// TIA Portal V21 export
FUNCTION_BLOCK "Mixed"   // FB1, LAD
BEGIN

REGION Network 1: Unknown part
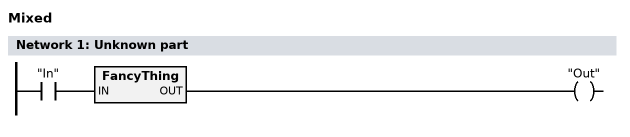
   // no SCL statement known for FancyThing: written as a call
   "Out" := FancyThing("In");
END_REGION

REGION Network 2 (SCL): SCL inside
END_REGION

REGION Network 3: Empty
END_REGION
END_FUNCTION_BLOCK
